TYPE "ST_SequenceStepDef"
VERSION : 0.1
   STRUCT
      StepNo : Int;
      Branch : Int;
      TimeClass : DInt;
      ExpectedTime : Time;
      StepName : String[120];
      AwaitingLabel : String[120];
      AwaitsPath : String[80];
   END_STRUCT;

END_TYPE

